(* IEC 61131-3 sources: volt/packages/volt-lsp-iec/test-corpus/awa-palletizer/Device/Plc Logic/Application/Library Manager/SysMem, 15 files *)

(* ---- SYSMEMALLOCAREA.pou ---- *)
FUNCTION SYSMEMALLOCAREA : POINTER TO BYTE
VAR_INPUT
	SZCOMPONENT : REFERENCE TO STRING;
	USTYPE : WORD;
	UDISIZE : __XWORD;
	PRESULT : POINTER TO RTS_IEC_RESULT;
END_VAR
END_FUNCTION

(* ---- SYSMEMALLOCCODE.pou ---- *)
FUNCTION SYSMEMALLOCCODE : POINTER TO BYTE
VAR_INPUT
	SZCOMPONENT : REFERENCE TO STRING;
	UDISIZE : __XWORD;
	PRESULT : POINTER TO RTS_IEC_RESULT;
END_VAR
END_FUNCTION

(* ---- SYSMEMALLOCDATA.pou ---- *)
FUNCTION SYSMEMALLOCDATA : POINTER TO BYTE
VAR_INPUT
	SZCOMPONENT : REFERENCE TO STRING;
	UDISIZE : __XWORD;
	PRESULT : POINTER TO RTS_IEC_RESULT;
END_VAR
END_FUNCTION

(* ---- SYSMEMCMP.pou ---- *)
FUNCTION SYSMEMCMP : DINT
VAR_INPUT
	PBUFFER1 : POINTER TO BYTE;
	PBUFFER2 : POINTER TO BYTE;
	UDICOUNT : __XWORD;
END_VAR
END_FUNCTION

(* ---- SYSMEMCPY.pou ---- *)
FUNCTION SYSMEMCPY : POINTER TO BYTE
VAR_INPUT
	PDEST : POINTER TO BYTE;
	PSRC : POINTER TO BYTE;
	UDICOUNT : __XWORD;
END_VAR
END_FUNCTION

(* ---- SYSMEMFORCESWAP.pou ---- *)
FUNCTION SYSMEMFORCESWAP : DINT
VAR_INPUT
	PBYBUFFER : POINTER TO BYTE;
	UDISIZE : UDINT;
	UDICOUNT : UDINT;
END_VAR
END_FUNCTION

(* ---- SYSMEMFREEAREA.pou ---- *)
FUNCTION SYSMEMFREEAREA : RTS_IEC_RESULT
VAR_INPUT
	SZCOMPONENT : REFERENCE TO STRING;
	PMEMORY : POINTER TO BYTE;
END_VAR
END_FUNCTION

(* ---- SYSMEMFREECODE.pou ---- *)
FUNCTION SYSMEMFREECODE : RTS_IEC_RESULT
VAR_INPUT
	SZCOMPONENT : REFERENCE TO STRING;
	PMEMORY : POINTER TO BYTE;
END_VAR
END_FUNCTION

(* ---- SYSMEMFREEDATA.pou ---- *)
FUNCTION SYSMEMFREEDATA : RTS_IEC_RESULT
VAR_INPUT
	SZCOMPONENT : REFERENCE TO STRING;
	PMEMORY : POINTER TO BYTE;
END_VAR
END_FUNCTION

(* ---- SYSMEMGETCURRENTHEAPSIZE.pou ---- *)
FUNCTION SYSMEMGETCURRENTHEAPSIZE : __XWORD
VAR_INPUT
	PRESULT : POINTER TO RTS_IEC_RESULT;
END_VAR
END_FUNCTION

(* ---- SYSMEMISVALIDPOINTER.pou ---- *)
FUNCTION SYSMEMISVALIDPOINTER : RTS_IEC_RESULT
VAR_INPUT
	PTR : POINTER TO BYTE;
	UDISIZE : __XWORD;
	BWRITE : BOOL;
END_VAR
END_FUNCTION

(* ---- SYSMEMMOVE.pou ---- *)
FUNCTION SYSMEMMOVE : POINTER TO BYTE
VAR_INPUT
	PDEST : POINTER TO BYTE;
	PSRC : POINTER TO BYTE;
	UDICOUNT : __XWORD;
END_VAR
END_FUNCTION

(* ---- SYSMEMREALLOCDATA.pou ---- *)
FUNCTION SYSMEMREALLOCDATA : POINTER TO BYTE
VAR_INPUT
	SZCOMPONENT : REFERENCE TO STRING;
	PMEMORY : POINTER TO BYTE;
	UDISIZE : __XWORD;
	PRESULT : POINTER TO RTS_IEC_RESULT;
END_VAR
END_FUNCTION

(* ---- SYSMEMSET.pou ---- *)
FUNCTION SYSMEMSET : POINTER TO BYTE
VAR_INPUT
	PDEST : POINTER TO BYTE;
	UDIVALUE : UDINT;
	UDICOUNT : __XWORD;
END_VAR
END_FUNCTION

(* ---- SYSMEMSWAP.pou ---- *)
FUNCTION SYSMEMSWAP : DINT
VAR_INPUT
	PBYBUFFER : POINTER TO BYTE;
	UDISIZE : UDINT;
	UDICOUNT : UDINT;
END_VAR
END_FUNCTION
